// TIA Portal V20 export
Screen "200APC1ayout"  1276x673
  ScreenItem "permanentareaborderrectangle" at 0,0 size 0x0  Type=HmiRectangle
  ScreenItem "Line_Header_X0_Y64" at 0,65 size 1276x0  Type=HmiLine
  ScreenItem "Button_Back" at 2,2 size 90x60  Type=HmiButton
  ScreenItem "Fusszeile_Button_ManualOPMode1_2" at 189,2 size 90x60  Type=HmiButton
  ScreenItem "Fusszeile_Button_ManualOPMode1_3" at 283,2 size 90x60  Type=HmiButton
  ScreenItem "面板容器_24" at 1092,4 size 88x58  Type=HmiFaceplateContainer
  ScreenItem "OPMode1_Blocked" at 1166,6 size 14x14  Type=HmiGraphicView
  ScreenItem "OPMode4_Foreground_Blocked" at 1092,4 size 88x58  Type=HmiGraphicView
  ScreenItem "Tec-Unit_LegendᆉY2" at 1184,2 size 90x60  Type=HmiButton
  ScreenItem "Fusszeile_Button_ManualOPMode1_1" at 95,2 size 90x60  Type=HmiButton
  ScreenItem "lOPMode1_4" at 991,3 size 90x60  Type=HmiButton
  ScreenItem "Graphic view_1" at 30,126 size 1170x343  Type=HmiGraphicView
  ScreenItem "Polygon_3" at 553,48 size 16x143  Type=HmiPolygon
  ScreenItem "Polygon_5" at 552,481 size 16x143  Type=HmiPolygon
  ScreenItem "Title_ScreenOverview_X390_Y2_2" at 459,513 size 201x23  Type=HmiTextBox
  ScreenItem "面板容器_8" at 220,212 size 59x49  Type=HmiFaceplateContainer
  ScreenItem "面板容器_1" at 214,313 size 61x49  Type=HmiFaceplateContainer
  ScreenItem "面板容器_3" at 8,209 size 146x52  Type=HmiFaceplateContainer
  ScreenItem "文本域_1" at 13,167 size 120x40  Type=HmiTextBox
  ScreenItem "面板容器_4" at 6,407 size 146x52  Type=HmiFaceplateContainer
  ScreenItem "文本域_2" at 6,364 size 120x40  Type=HmiTextBox
  ScreenItem "面板容器_5" at 1123,204 size 146x52  Type=HmiFaceplateContainer
  ScreenItem "面板容器_6" at 1125,403 size 146x52  Type=HmiFaceplateContainer
  ScreenItem "面板容器_10" at 1077,313 size 59x49  Type=HmiFaceplateContainer
  ScreenItem "面板容器_11" at 853,313 size 59x49  Type=HmiFaceplateContainer
  ScreenItem "面板容器_14" at 313,218 size 146x52  Type=HmiFaceplateContainer
  ScreenItem "文本域_7" at 310,176 size 120x40  Type=HmiTextBox
  ScreenItem "Rectangle TG1_1" at 13,577 size 234x81  Type=HmiRectangle
  ScreenItem "LED_1_Left_33" at 0,0 size 100x30  Type=HmiCircle
  ScreenItem "Text_DigitalOutputs_30" at 46,610 size 179x16  Type=HmiTextBox
  ScreenItem "Text_DigitalOutputs_1" at 46,634 size 179x16  Type=HmiTextBox
  ScreenItem "LED_1_Left_1" at 0,0 size 100x30  Type=HmiCircle
  ScreenItem "Text field Select Style" at 13,572 size 234x31  Type=HmiTextBox
  ScreenItem "文本域_18" at 200,191 size 100x20  Type=HmiTextBox
  ScreenItem "文本域_19" at 192,292 size 100x20  Type=HmiTextBox
  ScreenItem "文本域_20" at 832,292 size 100x20  Type=HmiTextBox
  ScreenItem "文本域_21" at 1040,292 size 100x20  Type=HmiTextBox
  ScreenItem "面板容器_16" at 568,619 size 146x52  Type=HmiFaceplateContainer
  ScreenItem "文本域_10" at 444,619 size 120x40  Type=HmiTextBox
  ScreenItem "面板容器_25" at 1113,562 size 146x52  Type=HmiFaceplateContainer
  ScreenItem "文本域_15" at 990,566 size 120x40  Type=HmiTextBox
  ScreenItem "文本域_16" at 990,623 size 120x40  Type=HmiTextBox
  ScreenItem "面板容器_22" at 1113,618 size 146x52  Type=HmiFaceplateContainer
  ScreenItem "文本域_17" at 714,619 size 120x40  Type=HmiTextBox
  ScreenItem "面板容器_23" at 837,619 size 146x52  Type=HmiFaceplateContainer
  ScreenItem "Title_ScreenOverview_X390_Y2_1" at 459,82 size 201x23  Type=HmiTextBox
  ScreenItem "Text_1" at 77,116 size 155x60  Type=HmiText
  ScreenItem "Text_2" at 958,116 size 205x60  Type=HmiText
  ScreenItem "文本域_5" at 8,70 size 120x40  Type=HmiTextBox
  ScreenItem "Title_ScreenOverview_X390_Y2_3" at 380,5 size 510x57  Type=HmiTextBox
  ScreenItem "按钮_2" at 300,70 size 140x60  Type=HmiButton
  ScreenItem "圆_9" at 0,0 size 100x30  Type=HmiCircle
  ScreenItem "按钮_1" at 300,502 size 140x60  Type=HmiButton
  ScreenItem "圆_1" at 0,0 size 100x30  Type=HmiCircle
  ScreenItem "按钮_4" at 677,502 size 140x60  Type=HmiButton
  ScreenItem "圆_3" at 0,0 size 100x30  Type=HmiCircle
  ScreenItem "按钮_5" at 837,502 size 140x60  Type=HmiButton
  ScreenItem "圆_4" at 0,0 size 100x30  Type=HmiCircle
  ScreenItem "文本域_6" at 1123,162 size 120x40  Type=HmiTextBox
  ScreenItem "文本域_8" at 1124,362 size 120x40  Type=HmiTextBox
  ScreenItem "文本域_9" at 280,352 size 120x40  Type=HmiTextBox
  ScreenItem "面板容器_2" at 280,392 size 146x52  Type=HmiFaceplateContainer
  ScreenItem "面板容器_7" at 428,392 size 146x52  Type=HmiFaceplateContainer
  ScreenItem "文本域_11" at 428,352 size 120x40  Type=HmiTextBox
  ScreenItem "面板容器_9" at 805,218 size 146x52  Type=HmiFaceplateContainer
  ScreenItem "文本域_12" at 805,177 size 120x40  Type=HmiTextBox
  ScreenItem "面板容器_12" at 978,474 size 146x52  Type=HmiFaceplateContainer
  ScreenItem "文本域_3" at 977,432 size 120x40  Type=HmiTextBox
  ScreenItem "面板容器_13" at 964,218 size 146x52  Type=HmiFaceplateContainer
  ScreenItem "文本域_13" at 960,177 size 120x40  Type=HmiTextBox
  ScreenItem "Rectangle_2" at 4,493 size 290x72  Type=HmiRectangle
  ScreenItem "Rectangle_3" at 8,474 size 284x41  Type=HmiRectangle
  ScreenItem "Text_11" at 4,476 size 288x41  Type=HmiText
  ScreenItem "Symbolic IO field_3" at 10,517 size 282x48  Type=HmiSymbolicIOField
  ScreenItem "Fusszeile_Button_ManualOPMode1_4" at 265,569 size 165x50  Type=HmiButton
